Fanuc KAREL source: KO00025.KL

PROGRAM KO00025
%NOLOCKGROUP
VAR
  P1: JOINTPOS
  P2: JOINTPOS
  P3: JOINTPOS
  OUT: POSITION
BEGIN
  OUT = FRAME(P1, P2, P3)
END KO00025
